(* IEC 61131-3 sources: Caravan/Archiv/12-04-19/Stations/Terminal/HMI/Network/Level_NET, 1 file *)

(* ---- ONE_Level_NET_Table.st ---- *)
#define OBJECTS_CONFIG

FUNCTION GLOBAL TAB ONE_Level_NET
-1$UINT, 0$UINT,
0$UINT, 0$UINT,

3$UDINT,
TO_UDINT(2980745877), "_MyIO", 0$UINT, 3$UINT, 0$UINT,
TO_UDINT(3621868871), "InputMyIO", 0$UINT, 0$UINT, 1$UINT,
TO_UDINT(2164406177), "Koordinates_Class", 0$UINT, 0$UINT, 1$UINT,

_NO_ATTR, TO_UDINT(1806949073), "INPUTMYIO1",

_NO_ATTR, TO_UDINT(579632894), "KOORDINATES_CLASS1",

//Internal connections
0$UDINT,
0$UDINT,
0$UDINT,
2$UDINT,
TO_UDINT(1), "Output_X_C", TO_UDINT(0), "sXDir",
TO_UDINT(1), "Output_Y_C", TO_UDINT(0), "sYDir",

//Initialization values
0$UDINT,
0$UDINT,

//Symbolic initialization values
0$UDINT,
0$UDINT,

//Initialization of string values
0$UDINT,
0$UDINT,

//Configuration of tasks (RealTime, Cyclic, Background)
0$UDINT,
0$UDINT,

0$UDINT,
1$UDINT,
TO_UDINT(1), (100)$UDINT, 4194303$DINT, 	//KOORDINATES_CLASS1

0$UDINT,
0$UDINT,

//External connections
0$UDINT,
1$UDINT,
TO_UDINT(0), "Lse", C_DIR, TO_UDINT(299963966), "Lse","Lse",

//Magic internal connections
0$UDINT,
0$UDINT,

//Configuration of timeslots of tasks (RealTime, Cyclic)
#ifdef __LSLLDR_TIMESLOTS__
0$UDINT,
0$UDINT,

0$UDINT,
0$UDINT,

#endif //__LSLLDR_TIMESLOTS__

//MultiMaster connections
#ifdef __LSLLDR_MULTIMASTER__
0$UDINT,
2$UDINT,
TO_UDINT(1), "Input_X_C", C_DIR, TO_UDINT(4258526131), "MachineControl.Level_Class1.Level_X_S",
TO_UDINT(1), "Input_Y_C", C_DIR, TO_UDINT(4229011844), "MachineControl.Level_Class1.Level_Y_S",
#endif //__LSLLDR_MULTIMASTER__

//Configuration for task ID (RealTime, CyclicTime)
#ifdef __LSLLDR_TASKID__
"\\\\TASKS2  "
0$UDINT,
0$UDINT,

0$UDINT,
1$UDINT,
(0)$UDINT, 	//KOORDINATES_CLASS1

0$UDINT,
0$UDINT,

#endif //__LSLLDR_TASKID__

END_FUNCTION
